(* IEC 61131-3 sources: avi-aoi-management/scripts/ai-eval/ngau-nhien/kho/st-ud10-thang-nang-2-tang/mau/src, 2 files *)

(* ---- KhoaDongCo.st ---- *)
FUNCTION_BLOCK KhoaDongCo
VAR_INPUT
    YC_LEN : BOOL;
    YC_XUONG : BOOL;
    CUA_DONG : BOOL;
    DUNG_KHAN : BOOL;
END_VAR
VAR_OUTPUT
    LEN : BOOL;
    XUONG : BOOL;
END_VAR
VAR
    choPhep : BOOL;
END_VAR
    choPhep := CUA_DONG AND NOT DUNG_KHAN AND NOT (YC_LEN AND YC_XUONG);
    LEN := YC_LEN AND choPhep;
    XUONG := YC_XUONG AND choPhep;
END_FUNCTION_BLOCK

(* ---- ThangNang2Tang.st ---- *)
FUNCTION_BLOCK ThangNang2Tang
VAR_INPUT
    GOI_1 : BOOL;
    GOI_2 : BOOL;
    CT_TANG_1 : BOOL;
    CT_TANG_2 : BOOL;
    CUA_DONG : BOOL;
    DUNG_KHAN : BOOL;
    RESET : BOOL;
    T_DI_CHUYEN : TIME;
END_VAR
VAR_OUTPUT
    LEN : BOOL;
    XUONG : BOOL;
    TRANG_THAI : INT;  (* 0 DUNG_YEN, 1 DI_LEN, 2 DI_XUONG, 9 LOI *)
    TANG : INT;        (* 0 chưa biết, 1, 2 *)
    MA_LOI : INT;      (* 0, 1 quá giờ, 2 dừng khẩn *)
END_VAR
VAR
    khoa : KhoaDongCo;
    tBuoc : TON;       (* ET = thời gian đã ở trạng thái hiện tại *)
    ttTruoc : INT;
END_VAR
    IF CT_TANG_1 AND NOT CT_TANG_2 THEN
        TANG := 1;
    ELSIF CT_TANG_2 AND NOT CT_TANG_1 THEN
        TANG := 2;
    END_IF
    tBuoc(IN := TRUE, PT := T#24h);

    IF DUNG_KHAN THEN
        TRANG_THAI := 9;
        MA_LOI := 2;
    ELSE
        CASE TRANG_THAI OF
        0:
            IF CUA_DONG AND NOT (GOI_1 AND GOI_2) THEN
                IF GOI_2 AND NOT CT_TANG_2 THEN
                    TRANG_THAI := 1;
                ELSIF GOI_1 AND NOT CT_TANG_1 THEN
                    TRANG_THAI := 2;
                END_IF
            END_IF
        1:
            IF CT_TANG_2 OR NOT CUA_DONG THEN
                TRANG_THAI := 0;
            ELSIF tBuoc.ET >= T_DI_CHUYEN THEN
                TRANG_THAI := 9;
                MA_LOI := 1;
            END_IF
        2:
            IF CT_TANG_1 OR NOT CUA_DONG THEN
                TRANG_THAI := 0;
            ELSIF tBuoc.ET >= T_DI_CHUYEN THEN
                TRANG_THAI := 9;
                MA_LOI := 1;
            END_IF
        9:
            IF RESET THEN
                TRANG_THAI := 0;
                MA_LOI := 0;
            END_IF
        END_CASE
    END_IF
    IF TRANG_THAI <> ttTruoc THEN
        tBuoc(IN := FALSE);
        tBuoc(IN := TRUE, PT := T#24h);
    END_IF
    ttTruoc := TRANG_THAI;

    khoa(YC_LEN := TRANG_THAI = 1, YC_XUONG := TRANG_THAI = 2, CUA_DONG := CUA_DONG, DUNG_KHAN := DUNG_KHAN);
    LEN := khoa.LEN;
    XUONG := khoa.XUONG;
END_FUNCTION_BLOCK
